Fanuc KAREL source: KT00879.KL

PROGRAM KT00879
%NOLOCKGROUP
VAR
  S1: STRING[80]
  S2: STRING[80]
  OUT: REAL
BEGIN
  S1 = 'A'
  S2 = 'B'
  S1 = 'A'
  S2 = 'B'
  OUT = TRUNC(S1)
END KT00879
